(* IEC 61131-3 sources: plcassist-cli/packages/volt-lsp-iec/test-corpus/CodesysTestProject/Device/Plc Logic/Application, 3 files *)

(* ---- VltFixtureCfc.fb ---- *)
FUNCTION_BLOCK VltFixtureCfc
VAR_INPUT
END_VAR
VAR_OUTPUT
END_VAR
VAR
END_VAR

(* @volt-graphical: CFC *)

END_FUNCTION_BLOCK

(* ---- VltFixtureSfc.fb ---- *)
FUNCTION_BLOCK VltFixtureSfc
VAR_INPUT
END_VAR
VAR_OUTPUT
END_VAR
VAR
END_VAR

(* @volt-graphical: SFC *)

END_FUNCTION_BLOCK

(* ---- PLC_PRG.prg ---- *)
PROGRAM PLC_PRG
VAR
END_VAR

END_PROGRAM
